// TIA Portal V21 export
// export: Created 2026-11-10T19:11:36.5902899Z, ExportSetting WithDefaults, DisplayName Totally Integrated Automation Portal, DisplayVersion V21 Update 3, DisplayName STEP 7 Professional, DisplayVersion V21 Update 3, DisplayName STEP 7 Safety, DisplayVersion V21, DisplayName Tech WebApplication, DisplayVersion V21, DisplayName WinCC Basic/Comfort/Advanced, DisplayVersion V21 Update 3, DisplayName WinCC Unified, DisplayVersion V21 Update 3
DATA_BLOCK "DB_Program_Alarm"   // DB21
// stored: AutoNumber true, DBAccessibleFromOPCUA true, DBAccessibleFromWebserver true, InstanceOfName Program_Alarm, OfSystemLibElement Program_Alarm, OfSystemLibVersion 1.0
"Program_Alarm"
   // // inherited from ALARM_BASE
   // VAR
   //    Alarm_ID : Event_ID;
   //    HANDLE : DWord;
   // END_VAR
   // VAR_INPUT
   //    SIG { ExternalWritable := 'False'} : Bool;
   //    TIMESTAMP { ExternalWritable := 'False'} : LDT;
   //    SD_1 : Variant;
   //    SD_2 : Variant;
   //    SD_3 : Variant;
   //    SD_4 : Variant;
   //    SD_5 : Variant;
   //    SD_6 : Variant;
   //    SD_7 : Variant;
   //    SD_8 : Variant;
   //    SD_9 : Variant;
   //    SD_10 : Variant;
   // END_VAR
   // VAR_OUTPUT
   //    Error { ExternalAccessible := 'False'; ExternalVisible := 'False'; ExternalWritable := 'False'} : Bool;
   //    Status { ExternalAccessible := 'False'; ExternalVisible := 'False'; ExternalWritable := 'False'} : Word;
   // END_VAR
   // VAR
   //    SD_0 { S7_SetPoint := 'True'} : AssocValue_0;
   // END_VAR
   // VAR RETAIN
   //    SIG_Edge_History { ExternalAccessible := 'False'; ExternalVisible := 'False'; ExternalWritable := 'False'} : Bool;
   // END_VAR
   // VAR
   //    INIT_FB_State : DWord;
   // END_VAR
BEGIN
END_DATA_BLOCK
